# EPICS substitutions: b-55B2VNC/src/main/c++/nds3-sdn/src/main/epics/ndssdnApp/Db/DeviceNDSSDNPUB.substitutions
##using the state machine in the device
#file "nds3_StateMachine.template" {
#	pattern
#	{	BOARDTYPE,
#		BOARDTYPEIDX,
#		CBS1,
#		CBS2,
#		STATEMACHINE_NAME
#	}
#	{	"SDN",
#		"0",
#		"TEST",
#		"FCT0",
#		"StateMachine"
#	}
#}

file "nds-sdn_pub.template" {
	pattern
	{	BOARDTYPE,
		BOARDTYPEIDX,
		CBS1,
		CBS2
	}
	{
		"SDN",
		"0",
		"TEST",
		"TEST",
	}
}
